Staubli VAL3: cycle_pause.pgx

public program cycle_pause()
begin
  rs:bToPause=true
  //  wait(rs:bIsPause==true)
  //  rs:bToPause=false
  //  logMsg("PLC:pausecycle")
end
